(* IEC 61131-3 sources: plc-ci-toolkit/tools/tests/fixtures/sample/src/Interfaces/I_Device, 1 file *)

(* ---- Start.method.decl.st ---- *)
METHOD Start
VAR_INPUT
    rSpeed_rpm : REAL;  // уставка скорости
END_VAR
